{attribute 'qualified_only'}
{attribute 'strict'}
TYPE E_Product_Type :
(
	Marinada := 0, Color
);
END_TYPE

(* stored: Version 1.1.0.1, ProductVersion 3.1.4024.12
   DUT E_Product_Type: Id {8e028360-d0d0-4a2e-af23-8948640999ef} *)
